PROGRAM MAIN
VAR
END_VAR

PRG_SafetyInterface();

END_PROGRAM

(* stored: Version 1.1.0.1
   POU MAIN: Id {6e8fa00b-7a4d-416c-8b1e-ef35aeb6bf5d}, SpecialFunc None *)
